(* Logix 5000 project; controller TFF vendor 1 type 14 code 107 rev 33.11; software revision 33.04; part 13 of 38 *)
(* tags used below, declared in another part *)
   AlarmAnalog : AlarmAnalog[50];   // Analog Alarm Array
   AlarmControl : AlarmControl;   // Alarm Control
   AlarmDeviation : AlarmDeviation[20];   // Control Loop Deviation Alarm Array
   AnalogPoint : AnalogInput[50];   // Analog Input Array
   BagInflate : BagInflate;
   CCPSystem : CCPSystem;   // CCP System Data
   ChartMark : ChartMark;   // Chart Mark
   Concentration : Concentration;
   ControlLoop : ControlLoop[20];   // Control Loop Array
   CriteriaFlag : CriteriaFlag;   // Criteria Flag used in CCP Recipe
   DerivedData : DerivedData;   // Derived data (user input and calculated values)
   Diafiltration : Diafiltration;
   DigitalOutput : BOOL[256];   // Digital Output Array these bits are sent to output cards.
   DigitalPoint : DigitalPoint[150];   // Digital Point Array
   Drive : Drive[11];   // Drives Array
   Exchange_OUT : Exchange_OUT;   // Exchange Outputs
   ExternalTCU : BOOL;   // Use of External TCU
   ExternalWeight : BOOL;   // Use of External Weight
   FlowPath : FlowPath[64];   // Flow Path Array
   FQ_Conc : ALIAS FOR Totalizer[0];   // Concentration Totalizer
   FQ_Diaf : ALIAS FOR Totalizer[1];   // DiafiltrationTotalizer
   Gateway : Gateway;   // Gateway Control
   LogVal : LoggedValue;   // Setpoints to be logged
   Membrane_Data : Membrane_Data;   // Membrane Data
   MiscBOOL : BOOL[64];   // Misc BOOL Values
   MiscDINT : DINT[32];   // Misc DINT Values
   MiscREAL : REAL[50];   // Misc Real Values
   Mixer : Mixer;   // Mixer config. structure
   Operation : Operation[6,251];   // Operation Table
   PCV101_Control : PCV_Control;   // PCV101 Control UDT
   PCV201_Control : PCV_Control;   // PCV201 Control UDT
   Phase : Phases[6];   // Phase Control Array
   Prompt : Prompt[7];   // Prompt Array
   PromptTimer : FBD_TIMER;   // Prompt Timer
   SysControl : SysControl;   // General system status and command
   TIC101Control : TCUControl;
   Timers : Timers[22];   // Timer Array
   Totalizer : Totalizers[20];   // Totalizers Array
   UserAlarm : UserAlarm;   // User Alarm (used in CCP Recipe)
   UserTotalizerManagement : UserTotalizerManagement;   // User Totalizer management
   Valve : Valve[100];   // Valve Array

        [2,19].AlarmTimerSP := 2, [2,19].AutoCloseTimer.ACC := 1007, [2,20].Tag := 'XV021', [2,20].CloseStatus := 1, [2,20].ZSOverride := 1, [2,20].EnableCfg := 1, [2,20].StatusWord := 4, [2,20].Status := 4, [2,20].OutputAddress := 52, [2,20].AlarmTimer.PRE := 2000, [2,20].AlarmTimerSP := 2, [2,20].AutoCloseTimer.ACC := 1004, [2,21].Tag := 'XV022', [2,21].Control := 1, [2,21].Auto := 1, [2,21].Manual := 1, [2,21].OpenStatus := 1, [2,21].ZSOverride := 1, [2,21].FailState := 1, [2,21].EnableCfg := 1, [2,21].StatusWord := 2, [2,21].Status := 2, [2,21].OutputAddress := 53, [2,21].AlarmTimer.PRE := 2000, [2,21].AlarmTimerSP := 2, [2,22].Tag := 'XV023', [2,22].CloseStatus := 1, [2,22].ZSOverride := 1, [2,22].EnableCfg := 1, [2,22].StatusWord := 4, [2,22].Status := 4, [2,22].OutputAddress := 54, [2,22].AlarmTimer.PRE := 2000, [2,22].AlarmTimerSP := 2, [2,22].AutoCloseTimer.ACC := 131, [2,23].Tag := 'XV024', [2,23].CloseStatus := 1, [2,23].ZSOverride := 1, [2,23].EnableCfg := 1, [2,23].StatusWord := 4, [2,23].Status := 4, [2,23].OutputAddress := 55, [2,23].AlarmTimer.PRE := 2000, [2,23].AlarmTimerSP := 2, [2,23].AutoCloseTimer.ACC := 1003, [2,24].Tag := 'XV025', [2,24].CloseStatus := 1, [2,24].ZSOverride := 1, [2,24].EnableCfg := 1, [2,24].StatusWord := 4, [2,24].Status := 4, [2,24].OutputAddress := 56, [2,24].AlarmTimer.PRE := 2000, [2,24].AlarmTimerSP := 2, [2,24].AutoCloseTimer.ACC := 1002, [2,25].Tag := 'XV026', [2,25].CloseStatus := 1, [2,25].ZSOverride := 1, [2,25].EnableCfg := 1, [2,25].StatusWord := 4,
        [2,25].Status := 4, [2,25].OutputAddress := 57, [2,25].AlarmTimer.PRE := 2000, [2,25].AlarmTimerSP := 2, [2,25].AutoCloseTimer.ACC := 1002, [2,26].Tag := 'XV028', [2,26].CloseStatus := 1, [2,26].ZSOverride := 1, [2,26].EnableCfg := 1, [2,26].StatusWord := 4, [2,26].Status := 4, [2,26].OutputAddress := 58, [2,26].AlarmTimer.PRE := 2000, [2,26].AlarmTimerSP := 2, [2,26].AutoCloseTimer.ACC := 1002, [2,27].Tag := 'XV029', [2,27].CloseStatus := 1, [2,27].ZSOverride := 1, [2,27].EnableCfg := 1, [2,27].StatusWord := 4, [2,27].Status := 4, [2,27].OutputAddress := 59, [2,27].AlarmTimer.PRE := 2000, [2,27].AlarmTimerSP := 2, [2,28].Tag := 'XV030', [2,28].CloseStatus := 1, [2,28].ZSOverride := 1, [2,28].EnableCfg := 1, [2,28].StatusWord := 4, [2,28].Status := 4, [2,28].OutputAddress := 60, [2,28].AlarmTimer.PRE := 2000, [2,28].AlarmTimerSP := 2, [2,29].Tag := 'XV031', [2,29].Control := 1, [2,29].Auto := 1, [2,29].Manual := 1, [2,29].OpenStatus := 1, [2,29].ZSOverride := 1, [2,29].FailState := 1, [2,29].EnableCfg := 1, [2,29].StatusWord := 2, [2,29].Status := 2, [2,29].OutputAddress := 61, [2,29].AlarmTimer.PRE := 2000, [2,29].AlarmTimerSP := 2, [2,29].AutoCloseTimer.ACC := 1068, [2,30].Tag := 'XV033', [2,30].CloseStatus := 1, [2,30].ZSOverride := 1, [2,30].EnableCfg := 1, [2,30].StatusWord := 4, [2,30].Status := 4, [2,30].OutputAddress := 62, [2,30].AlarmTimer.PRE := 2000, [2,30].AlarmTimerSP := 2, [2,30].AutoCloseTimer.ACC := 1069, [2,31].Tag := 'XV034', [2,31].CloseStatus := 1, [2,31].ZSOverride := 1,
        [2,31].EnableCfg := 1, [2,31].StatusWord := 4, [2,31].Status := 4, [2,31].OutputAddress := 63, [2,31].AlarmTimer.PRE := 2000, [2,31].AlarmTimerSP := 2, [2,31].AutoCloseTimer.ACC := 131, [2,32].CloseStatus := 1, [2,32].PriorityCfg := 1, [2,32].ZSOpenAddress := 32, [2,32].OutputAddress := 68, [2,32].AlarmTimer.PRE := 2000, [2,32].AlarmTimerSP := 2, [2,32].AutoCloseTimer.ACC := 1059, [2,33].OpenStatus := 1, [2,33].PriorityCfg := 1, [2,33].FailState := 1, [2,33].ZSCloseAddress := 33, [2,33].OutputAddress := 69, [2,33].AlarmTimer.PRE := 2000, [2,33].AlarmTimerSP := 2, [2,33].AutoCloseTimer.ACC := 1123, [2,34].OpenStatus := 1, [2,34].PriorityCfg := 1, [2,34].FailState := 1, [2,34].ZSCloseAddress := 34, [2,34].OutputAddress := 70, [2,34].AlarmTimer.PRE := 2000, [2,34].AlarmTimerSP := 2, [2,34].AutoCloseTimer.ACC := 1095, [2,35].OpenStatus := 1, [2,35].PriorityCfg := 1, [2,35].FailState := 1, [2,35].ZSCloseAddress := 35, [2,35].OutputAddress := 71, [2,35].AlarmTimer.PRE := 2000, [2,35].AlarmTimerSP := 2, [2,35].AutoCloseTimer.ACC := 1127, [2,36].OpenStatus := 1, [2,36].PriorityCfg := 1, [2,36].FailState := 1, [2,36].ZSCloseAddress := 36, [2,36].OutputAddress := 72, [2,36].AlarmTimer.PRE := 2000, [2,36].AlarmTimerSP := 2, [2,36].AutoCloseTimer.ACC := 1004, [2,37].CloseStatus := 1, [2,37].PriorityCfg := 1, [2,37].ZSOpenAddress := 37, [2,37].OutputAddress := 73, [2,37].AlarmTimer.PRE := 2000, [2,37].AlarmTimerSP := 2, [2,37].AutoCloseTimer.ACC := 1121, [2,38].CloseStatus := 1, [2,38].Priority := 1, [2,38].PriorityCfg := 1, [2,38].ZSOpenAddress := 38, [2,38].OutputAddress := 40, [2,38].AlarmTimer.PRE := 2000, [2,38].AlarmTimerSP := 2,
        [2,38].AutoCloseTimer.ACC := 1135, [2,39].CloseStatus := 1, [2,39].Priority := 1, [2,39].PriorityCfg := 1, [2,39].ZSOpenAddress := 39, [2,39].OutputAddress := 41, [2,39].AlarmTimer.PRE := 2000, [2,39].AlarmTimerSP := 2, [2,39].AutoCloseTimer.ACC := 1121, [2,40].CloseStatus := 1, [2,40].Priority := 1, [2,40].PriorityCfg := 1, [2,40].ZSOpenAddress := 40, [2,40].OutputAddress := 42, [2,40].AlarmTimer.PRE := 2000, [2,40].AlarmTimerSP := 2, [2,40].AutoCloseTimer.ACC := 1112, [2,41].CloseStatus := 1, [2,41].Priority := 1, [2,41].PriorityCfg := 1, [2,41].ZSOpenAddress := 41, [2,41].OutputAddress := 43, [2,41].AlarmTimer.PRE := 2000, [2,41].AlarmTimerSP := 2, [2,42].CloseStatus := 1, [2,42].Priority := 1, [2,42].PriorityCfg := 1, [2,42].ZSOpenAddress := 42, [2,42].OutputAddress := 44, [2,42].AlarmTimer.PRE := 2000, [2,42].AlarmTimerSP := 2, [2,43].CloseStatus := 1, [2,43].Priority := 1, [2,43].PriorityCfg := 1, [2,43].ZSOpenAddress := 43, [2,43].OutputAddress := 52, [2,43].AlarmTimer.PRE := 2000, [2,43].AlarmTimerSP := 2, [2,44].CloseStatus := 1, [2,44].Priority := 1, [2,44].PriorityCfg := 1, [2,44].ZSOpenAddress := 44, [2,44].OutputAddress := 53, [2,44].AlarmTimer.PRE := 2000, [2,44].AlarmTimerSP := 2, [2,45].CloseStatus := 1, [2,45].Priority := 1, [2,45].PriorityCfg := 1, [2,45].ZSOpenAddress := 45, [2,45].OutputAddress := 54, [2,45].AlarmTimer.PRE := 2000, [2,45].AlarmTimerSP := 2, [2,46].CloseStatus := 1, [2,46].Priority := 1, [2,46].PriorityCfg := 1, [2,46].ZSOpenAddress := 46, [2,46].OutputAddress := 55, [2,46].AlarmTimer.PRE := 2000, [2,46].AlarmTimerSP := 2, [2,47].OpenStatus := 1,
        [2,47].Priority := 1, [2,47].PriorityCfg := 1, [2,47].FailState := 1, [2,47].ZSCloseAddress := 47, [2,47].OutputAddress := 45, [2,47].AlarmTimer.PRE := 2000, [2,47].AlarmTimerSP := 2, [2,48].FailState := 1, [2,48].ZSCloseAddress := 48, [2,48].OutputAddress := 80, [2,49].FailState := 1, [2,49].ZSCloseAddress := 49, [2,49].OutputAddress := 81, [2,50].FailState := 1, [2,50].ZSCloseAddress := 50, [2,50].OutputAddress := 82, [2,51].OpenStatus := 1, [2,51].FailState := 1, [2,51].ZSCloseAddress := 51, [2,51].OutputAddress := 83, [2,52].OpenStatus := 1, [2,52].FailState := 1, [2,52].ZSCloseAddress := 52, [2,52].OutputAddress := 84, [2,53].CloseStatus := 1, [2,53].FailState := 1, [2,53].ZSCloseAddress := 53, [2,53].OutputAddress := 85, [2,54].CloseStatus := 1, [2,54].FailState := 1, [2,54].ZSCloseAddress := 54, [2,54].OutputAddress := 86, [2,55].CloseStatus := 1, [2,55].FailState := 1, [2,55].ZSCloseAddress := 55, [2,55].OutputAddress := 87, [2,56].CloseStatus := 1, [2,58].CloseStatus := 1, [2,59].CloseStatus := 1, [3,0].CloseStatus := 1, [3,0].EnableCfg := 1, [3,0].StatusWord := 4, [3,0].Status := 4, [3,0].OutputAddress := 32, [3,1].CloseStatus := 1, [3,1].EnableCfg := 1, [3,1].StatusWord := 4, [3,1].Status := 4, [3,1].OutputAddress := 33, [3,2].CloseStatus := 1, [3,2].EnableCfg := 1, [3,2].StatusWord := 4, [3,2].Status := 4, [3,2].OutputAddress := 34, [3,3].CloseStatus := 1, [3,3].EnableCfg := 1, [3,3].StatusWord := 4, [3,3].Status := 4, [3,3].OutputAddress := 35, [3,4].CloseStatus := 1,
        [3,4].EnableCfg := 1, [3,4].StatusWord := 4, [3,4].Status := 4, [3,4].OutputAddress := 36, [3,5].CloseStatus := 1, [3,5].EnableCfg := 1, [3,5].StatusWord := 4, [3,5].Status := 4, [3,5].OutputAddress := 37, [3,6].CloseStatus := 1, [3,6].EnableCfg := 1, [3,6].StatusWord := 4, [3,6].Status := 4, [3,6].OutputAddress := 38, [3,7].CloseStatus := 1, [3,7].EnableCfg := 1, [3,7].StatusWord := 4, [3,7].Status := 4, [3,7].OutputAddress := 39, [3,8].CloseStatus := 1, [3,8].EnableCfg := 1, [3,8].StatusWord := 4, [3,8].Status := 4, [3,8].OutputAddress := 40, [3,9].CloseStatus := 1, [3,9].EnableCfg := 1, [3,9].StatusWord := 4, [3,9].Status := 4, [3,9].OutputAddress := 41, [3,10].CloseStatus := 1, [3,10].EnableCfg := 1, [3,10].StatusWord := 4, [3,10].Status := 4, [3,10].OutputAddress := 42, [3,11].CloseStatus := 1, [3,11].FailState := 1, [3,11].EnableCfg := 1, [3,11].StatusWord := 4, [3,11].Status := 4, [3,11].OutputAddress := 43, [3,12].CloseStatus := 1, [3,12].FailState := 1, [3,12].EnableCfg := 1, [3,12].StatusWord := 4, [3,12].Status := 4, [3,12].OutputAddress := 44, [3,13].CloseStatus := 1, [3,13].FailState := 1, [3,13].EnableCfg := 1, [3,13].StatusWord := 4, [3,13].Status := 4, [3,13].OutputAddress := 45, [3,14].CloseStatus := 1, [3,14].EnableCfg := 1, [3,14].StatusWord := 4, [3,14].Status := 4, [3,14].OutputAddress := 46, [3,15].CloseStatus := 1, [3,15].FailState := 1, [3,15].EnableCfg := 1,
        [3,15].StatusWord := 4, [3,15].Status := 4, [3,15].OutputAddress := 47, [3,16].CloseStatus := 1, [3,16].EnableCfg := 1, [3,16].StatusWord := 4, [3,16].Status := 4, [3,16].OutputAddress := 48, [3,17].CloseStatus := 1, [3,17].FailState := 1, [3,17].EnableCfg := 1, [3,17].StatusWord := 4, [3,17].Status := 4, [3,17].OutputAddress := 49, [3,18].CloseStatus := 1, [3,18].EnableCfg := 1, [3,18].StatusWord := 4, [3,18].Status := 4, [3,18].OutputAddress := 50, [3,19].CloseStatus := 1, [3,19].EnableCfg := 1, [3,19].StatusWord := 4, [3,19].Status := 4, [3,19].OutputAddress := 51, [3,20].CloseStatus := 1, [3,20].EnableCfg := 1, [3,20].StatusWord := 4, [3,20].Status := 4, [3,20].OutputAddress := 52, [3,21].CloseStatus := 1, [3,21].FailState := 1, [3,21].EnableCfg := 1, [3,21].StatusWord := 4, [3,21].Status := 4, [3,21].OutputAddress := 53, [3,22].CloseStatus := 1, [3,22].EnableCfg := 1, [3,22].StatusWord := 4, [3,22].Status := 4, [3,22].OutputAddress := 54, [3,23].CloseStatus := 1, [3,23].EnableCfg := 1, [3,23].StatusWord := 4, [3,23].Status := 4, [3,23].OutputAddress := 55, [3,24].CloseStatus := 1, [3,24].EnableCfg := 1, [3,24].StatusWord := 4, [3,24].Status := 4, [3,24].OutputAddress := 56, [3,25].CloseStatus := 1, [3,25].EnableCfg := 1, [3,25].StatusWord := 4, [3,25].Status := 4, [3,25].OutputAddress := 57, [3,26].CloseStatus := 1, [3,26].EnableCfg := 1, [3,26].StatusWord := 4, [3,26].Status := 4, [3,26].OutputAddress := 58,
        [3,27].CloseStatus := 1, [3,27].EnableCfg := 1, [3,27].StatusWord := 4, [3,27].Status := 4, [3,27].OutputAddress := 59, [3,28].CloseStatus := 1, [3,28].EnableCfg := 1, [3,28].StatusWord := 4, [3,28].Status := 4, [3,28].OutputAddress := 60, [3,29].CloseStatus := 1, [3,29].FailState := 1, [3,29].EnableCfg := 1, [3,29].StatusWord := 4, [3,29].Status := 4, [3,29].OutputAddress := 61, [3,30].CloseStatus := 1, [3,30].EnableCfg := 1, [3,30].StatusWord := 4, [3,30].Status := 4, [3,30].OutputAddress := 62, [3,31].CloseStatus := 1, [3,31].EnableCfg := 1, [3,31].StatusWord := 4, [3,31].Status := 4, [3,31].OutputAddress := 63, [4,0].Tag := 'XV001', [4,0].CloseStatus := 1, [4,0].ZSOverride := 1, [4,0].EnableCfg := 1, [4,0].StatusWord := 4, [4,0].Status := 4, [4,0].OutputAddress := 32, [4,0].AlarmTimer.PRE := 2000, [4,0].AlarmTimerSP := 2, [4,1].Tag := 'XV002', [4,1].CloseStatus := 1, [4,1].ZSOverride := 1, [4,1].EnableCfg := 1, [4,1].StatusWord := 4, [4,1].Status := 4, [4,1].OutputAddress := 33, [4,1].AlarmTimer.PRE := 2000, [4,1].AlarmTimerSP := 2, [4,1].AutoCloseTimer.ACC := 1103, [4,2].Tag := 'XV003', [4,2].CloseStatus := 1, [4,2].ZSOverride := 1, [4,2].EnableCfg := 1, [4,2].StatusWord := 4, [4,2].Status := 4, [4,2].OutputAddress := 34, [4,2].AlarmTimer.PRE := 2000, [4,2].AlarmTimerSP := 2, [4,2].AutoCloseTimer.ACC := 1032, [4,3].Tag := 'XV004', [4,3].CloseStatus := 1, [4,3].ZSOverride := 1, [4,3].EnableCfg := 1, [4,3].StatusWord := 4,
        [4,3].Status := 4, [4,3].OutputAddress := 35, [4,3].AlarmTimer.PRE := 2000, [4,3].AlarmTimerSP := 2, [4,3].AutoCloseTimer.ACC := 1115, [4,4].Tag := 'XV005', [4,4].CloseStatus := 1, [4,4].ZSOverride := 1, [4,4].EnableCfg := 1, [4,4].StatusWord := 4, [4,4].Status := 4, [4,4].OutputAddress := 36, [4,4].AlarmTimer.PRE := 2000, [4,4].AlarmTimerSP := 2, [4,4].AutoCloseTimer.ACC := 1104, [4,5].Tag := 'XV006', [4,5].CloseStatus := 1, [4,5].ZSOverride := 1, [4,5].EnableCfg := 1, [4,5].StatusWord := 4, [4,5].Status := 4, [4,5].OutputAddress := 37, [4,5].AlarmTimer.PRE := 2000, [4,5].AlarmTimerSP := 2, [4,5].AutoCloseTimer.ACC := 1104, [4,6].Tag := 'XV007', [4,6].CloseStatus := 1, [4,6].ZSOverride := 1, [4,6].EnableCfg := 1, [4,6].StatusWord := 4, [4,6].Status := 4, [4,6].OutputAddress := 38, [4,6].AlarmTimer.PRE := 2000, [4,6].AlarmTimerSP := 2, [4,6].AutoCloseTimer.ACC := 1104, [4,7].Tag := 'XV008', [4,7].CloseStatus := 1, [4,7].ZSOverride := 1, [4,7].EnableCfg := 1, [4,7].StatusWord := 4, [4,7].Status := 4, [4,7].OutputAddress := 39, [4,7].AlarmTimer.PRE := 2000, [4,7].AlarmTimerSP := 2, [4,7].AutoCloseTimer.ACC := 1104, [4,8].Tag := 'XV009', [4,8].CloseStatus := 1, [4,8].ZSOverride := 1, [4,8].EnableCfg := 1, [4,8].StatusWord := 4, [4,8].Status := 4, [4,8].OutputAddress := 40, [4,8].AlarmTimer.PRE := 2000, [4,8].AlarmTimerSP := 2, [4,8].AutoCloseTimer.ACC := 1104, [4,9].Tag := 'XV010', [4,9].CloseStatus := 1, [4,9].ZSOverride := 1, [4,9].EnableCfg := 1, [4,9].StatusWord := 4,
        [4,9].Status := 4, [4,9].OutputAddress := 41, [4,9].AlarmTimer.PRE := 2000, [4,9].AlarmTimerSP := 2, [4,9].AutoCloseTimer.ACC := 1105, [4,10].Tag := 'XV011', [4,10].CloseStatus := 1, [4,10].ZSOverride := 1, [4,10].EnableCfg := 1, [4,10].StatusWord := 4, [4,10].Status := 4, [4,10].OutputAddress := 42, [4,10].AlarmTimer.PRE := 2000, [4,10].AlarmTimerSP := 2, [4,10].AutoCloseTimer.ACC := 1104, [4,11].Tag := 'XV012', [4,11].Control := 1, [4,11].Auto := 1, [4,11].Manual := 1, [4,11].OpenStatus := 1, [4,11].ZSOverride := 1, [4,11].FailState := 1, [4,11].EnableCfg := 1, [4,11].StatusWord := 2, [4,11].Status := 2, [4,11].OutputAddress := 43, [4,11].AlarmTimer.PRE := 2000, [4,11].AlarmTimerSP := 2, [4,11].AutoCloseTimer.ACC := 1103, [4,12].Tag := 'XV013', [4,12].Control := 1, [4,12].Auto := 1, [4,12].Manual := 1, [4,12].OpenStatus := 1, [4,12].ZSOverride := 1, [4,12].FailState := 1, [4,12].EnableCfg := 1, [4,12].StatusWord := 2, [4,12].Status := 2, [4,12].OutputAddress := 44, [4,12].AlarmTimer.PRE := 2000, [4,12].AlarmTimerSP := 2, [4,12].AutoCloseTimer.ACC := 1072, [4,13].Tag := 'XV014', [4,13].Control := 1, [4,13].Auto := 1, [4,13].Manual := 1, [4,13].OpenStatus := 1, [4,13].ZSOverride := 1, [4,13].FailState := 1, [4,13].EnableCfg := 1, [4,13].StatusWord := 2, [4,13].Status := 2, [4,13].OutputAddress := 45, [4,13].AlarmTimer.PRE := 2000, [4,13].AlarmTimerSP := 2, [4,13].AutoCloseTimer.ACC := 1016, [4,14].Tag := 'XV015', [4,14].CloseStatus := 1, [4,14].ZSOverride := 1,
        [4,14].EnableCfg := 1, [4,14].StatusWord := 4, [4,14].Status := 4, [4,14].OutputAddress := 46, [4,14].AlarmTimer.PRE := 2000, [4,14].AlarmTimerSP := 2, [4,15].Tag := 'XV016', [4,15].Control := 1, [4,15].Auto := 1, [4,15].Manual := 1, [4,15].OpenStatus := 1, [4,15].ZSOverride := 1, [4,15].FailState := 1, [4,15].EnableCfg := 1, [4,15].StatusWord := 2, [4,15].Status := 2, [4,15].OutputAddress := 47, [4,15].AlarmTimer.PRE := 2000, [4,15].AlarmTimerSP := 2, [4,16].Tag := 'XV017', [4,16].CloseStatus := 1, [4,16].ZSOverride := 1, [4,16].EnableCfg := 1, [4,16].StatusWord := 4, [4,16].Status := 4, [4,16].OutputAddress := 48, [4,16].AlarmTimer.PRE := 2000, [4,16].AlarmTimerSP := 2, [4,17].Tag := 'XV018', [4,17].Control := 1, [4,17].Auto := 1, [4,17].Manual := 1, [4,17].OpenStatus := 1, [4,17].ZSOverride := 1, [4,17].FailState := 1, [4,17].EnableCfg := 1, [4,17].StatusWord := 2, [4,17].Status := 2, [4,17].OutputAddress := 49, [4,17].AlarmTimer.PRE := 2000, [4,17].AlarmTimerSP := 2, [4,17].AutoCloseTimer.ACC := 1594, [4,18].Tag := 'XV019', [4,18].CloseStatus := 1, [4,18].ZSOverride := 1, [4,18].EnableCfg := 1, [4,18].StatusWord := 4, [4,18].Status := 4, [4,18].OutputAddress := 50, [4,18].AlarmTimer.PRE := 2000, [4,18].AlarmTimerSP := 2, [4,18].AutoCloseTimer.ACC := 137, [4,19].Tag := 'XV020', [4,19].CloseStatus := 1, [4,19].ZSOverride := 1, [4,19].EnableCfg := 1, [4,19].StatusWord := 4, [4,19].Status := 4, [4,19].OutputAddress := 51, [4,19].AlarmTimer.PRE := 2000,
        [4,19].AlarmTimerSP := 2, [4,19].AutoCloseTimer.ACC := 1007, [4,20].Tag := 'XV021', [4,20].CloseStatus := 1, [4,20].ZSOverride := 1, [4,20].EnableCfg := 1, [4,20].StatusWord := 4, [4,20].Status := 4, [4,20].OutputAddress := 52, [4,20].AlarmTimer.PRE := 2000, [4,20].AlarmTimerSP := 2, [4,20].AutoCloseTimer.ACC := 1004, [4,21].Tag := 'XV022', [4,21].Control := 1, [4,21].Auto := 1, [4,21].Manual := 1, [4,21].OpenStatus := 1, [4,21].ZSOverride := 1, [4,21].FailState := 1, [4,21].EnableCfg := 1, [4,21].StatusWord := 2, [4,21].Status := 2, [4,21].OutputAddress := 53, [4,21].AlarmTimer.PRE := 2000, [4,21].AlarmTimerSP := 2, [4,22].Tag := 'XV023', [4,22].CloseStatus := 1, [4,22].ZSOverride := 1, [4,22].EnableCfg := 1, [4,22].StatusWord := 4, [4,22].Status := 4, [4,22].OutputAddress := 54, [4,22].AlarmTimer.PRE := 2000, [4,22].AlarmTimerSP := 2, [4,22].AutoCloseTimer.ACC := 131, [4,23].Tag := 'XV024', [4,23].CloseStatus := 1, [4,23].ZSOverride := 1, [4,23].EnableCfg := 1, [4,23].StatusWord := 4, [4,23].Status := 4, [4,23].OutputAddress := 55, [4,23].AlarmTimer.PRE := 2000, [4,23].AlarmTimerSP := 2, [4,23].AutoCloseTimer.ACC := 1003, [4,24].Tag := 'XV025', [4,24].CloseStatus := 1, [4,24].ZSOverride := 1, [4,24].EnableCfg := 1, [4,24].StatusWord := 4, [4,24].Status := 4, [4,24].OutputAddress := 56, [4,24].AlarmTimer.PRE := 2000, [4,24].AlarmTimerSP := 2, [4,24].AutoCloseTimer.ACC := 1002, [4,25].Tag := 'XV026', [4,25].CloseStatus := 1, [4,25].ZSOverride := 1, [4,25].EnableCfg := 1, [4,25].StatusWord := 4,
        [4,25].Status := 4, [4,25].OutputAddress := 57, [4,25].AlarmTimer.PRE := 2000, [4,25].AlarmTimerSP := 2, [4,25].AutoCloseTimer.ACC := 1002, [4,26].Tag := 'XV028', [4,26].CloseStatus := 1, [4,26].ZSOverride := 1, [4,26].EnableCfg := 1, [4,26].StatusWord := 4, [4,26].Status := 4, [4,26].OutputAddress := 58, [4,26].AlarmTimer.PRE := 2000, [4,26].AlarmTimerSP := 2, [4,26].AutoCloseTimer.ACC := 1002, [4,27].Tag := 'XV029', [4,27].CloseStatus := 1, [4,27].ZSOverride := 1, [4,27].EnableCfg := 1, [4,27].StatusWord := 4, [4,27].Status := 4, [4,27].OutputAddress := 59, [4,27].AlarmTimer.PRE := 2000, [4,27].AlarmTimerSP := 2, [4,28].Tag := 'XV030', [4,28].CloseStatus := 1, [4,28].ZSOverride := 1, [4,28].EnableCfg := 1, [4,28].StatusWord := 4, [4,28].Status := 4, [4,28].OutputAddress := 60, [4,28].AlarmTimer.PRE := 2000, [4,28].AlarmTimerSP := 2, [4,29].Tag := 'XV031', [4,29].Control := 1, [4,29].Auto := 1, [4,29].Manual := 1, [4,29].OpenStatus := 1, [4,29].ZSOverride := 1, [4,29].FailState := 1, [4,29].EnableCfg := 1, [4,29].StatusWord := 2, [4,29].Status := 2, [4,29].OutputAddress := 61, [4,29].AlarmTimer.PRE := 2000, [4,29].AlarmTimerSP := 2, [4,29].AutoCloseTimer.ACC := 1068, [4,30].Tag := 'XV033', [4,30].CloseStatus := 1, [4,30].ZSOverride := 1, [4,30].EnableCfg := 1, [4,30].StatusWord := 4, [4,30].Status := 4, [4,30].OutputAddress := 62, [4,30].AlarmTimer.PRE := 2000, [4,30].AlarmTimerSP := 2, [4,30].AutoCloseTimer.ACC := 1069, [4,31].Tag := 'XV034', [4,31].CloseStatus := 1, [4,31].ZSOverride := 1,
        [4,31].EnableCfg := 1, [4,31].StatusWord := 4, [4,31].Status := 4, [4,31].OutputAddress := 63, [4,31].AlarmTimer.PRE := 2000, [4,31].AlarmTimerSP := 2, [4,31].AutoCloseTimer.ACC := 131, [4,32].CloseStatus := 1, [4,32].PriorityCfg := 1, [4,32].ZSOpenAddress := 32, [4,32].OutputAddress := 68, [4,32].AlarmTimer.PRE := 2000, [4,32].AlarmTimerSP := 2, [4,32].AutoCloseTimer.ACC := 1059, [4,33].OpenStatus := 1, [4,33].PriorityCfg := 1, [4,33].FailState := 1, [4,33].ZSCloseAddress := 33, [4,33].OutputAddress := 69, [4,33].AlarmTimer.PRE := 2000, [4,33].AlarmTimerSP := 2, [4,33].AutoCloseTimer.ACC := 1123, [4,34].OpenStatus := 1, [4,34].PriorityCfg := 1, [4,34].FailState := 1, [4,34].ZSCloseAddress := 34, [4,34].OutputAddress := 70, [4,34].AlarmTimer.PRE := 2000, [4,34].AlarmTimerSP := 2, [4,34].AutoCloseTimer.ACC := 1095, [4,35].OpenStatus := 1, [4,35].PriorityCfg := 1, [4,35].FailState := 1, [4,35].ZSCloseAddress := 35, [4,35].OutputAddress := 71, [4,35].AlarmTimer.PRE := 2000, [4,35].AlarmTimerSP := 2, [4,35].AutoCloseTimer.ACC := 1127, [4,36].OpenStatus := 1, [4,36].PriorityCfg := 1, [4,36].FailState := 1, [4,36].ZSCloseAddress := 36, [4,36].OutputAddress := 72, [4,36].AlarmTimer.PRE := 2000, [4,36].AlarmTimerSP := 2, [4,36].AutoCloseTimer.ACC := 1004, [4,37].CloseStatus := 1, [4,37].PriorityCfg := 1, [4,37].ZSOpenAddress := 37, [4,37].OutputAddress := 73, [4,37].AlarmTimer.PRE := 2000, [4,37].AlarmTimerSP := 2, [4,37].AutoCloseTimer.ACC := 1121, [4,38].CloseStatus := 1, [4,38].Priority := 1, [4,38].PriorityCfg := 1, [4,38].ZSOpenAddress := 38, [4,38].OutputAddress := 40, [4,38].AlarmTimer.PRE := 2000, [4,38].AlarmTimerSP := 2,
        [4,38].AutoCloseTimer.ACC := 1135, [4,39].CloseStatus := 1, [4,39].Priority := 1, [4,39].PriorityCfg := 1, [4,39].ZSOpenAddress := 39, [4,39].OutputAddress := 41, [4,39].AlarmTimer.PRE := 2000, [4,39].AlarmTimerSP := 2, [4,39].AutoCloseTimer.ACC := 1121, [4,40].CloseStatus := 1, [4,40].Priority := 1, [4,40].PriorityCfg := 1, [4,40].ZSOpenAddress := 40, [4,40].OutputAddress := 42, [4,40].AlarmTimer.PRE := 2000, [4,40].AlarmTimerSP := 2, [4,40].AutoCloseTimer.ACC := 1112, [4,41].CloseStatus := 1, [4,41].Priority := 1, [4,41].PriorityCfg := 1, [4,41].ZSOpenAddress := 41, [4,41].OutputAddress := 43, [4,41].AlarmTimer.PRE := 2000, [4,41].AlarmTimerSP := 2, [4,42].CloseStatus := 1, [4,42].Priority := 1, [4,42].PriorityCfg := 1, [4,42].ZSOpenAddress := 42, [4,42].OutputAddress := 44, [4,42].AlarmTimer.PRE := 2000, [4,42].AlarmTimerSP := 2, [4,43].CloseStatus := 1, [4,43].Priority := 1, [4,43].PriorityCfg := 1, [4,43].ZSOpenAddress := 43, [4,43].OutputAddress := 52, [4,43].AlarmTimer.PRE := 2000, [4,43].AlarmTimerSP := 2, [4,44].CloseStatus := 1, [4,44].Priority := 1, [4,44].PriorityCfg := 1, [4,44].ZSOpenAddress := 44, [4,44].OutputAddress := 53, [4,44].AlarmTimer.PRE := 2000, [4,44].AlarmTimerSP := 2, [4,45].CloseStatus := 1, [4,45].Priority := 1, [4,45].PriorityCfg := 1, [4,45].ZSOpenAddress := 45, [4,45].OutputAddress := 54, [4,45].AlarmTimer.PRE := 2000, [4,45].AlarmTimerSP := 2, [4,46].CloseStatus := 1, [4,46].Priority := 1, [4,46].PriorityCfg := 1, [4,46].ZSOpenAddress := 46, [4,46].OutputAddress := 55, [4,46].AlarmTimer.PRE := 2000, [4,46].AlarmTimerSP := 2, [4,47].OpenStatus := 1,
        [4,47].Priority := 1, [4,47].PriorityCfg := 1, [4,47].FailState := 1, [4,47].ZSCloseAddress := 47, [4,47].OutputAddress := 45, [4,47].AlarmTimer.PRE := 2000, [4,47].AlarmTimerSP := 2, [4,48].FailState := 1, [4,48].ZSCloseAddress := 48, [4,48].OutputAddress := 80, [4,49].FailState := 1, [4,49].ZSCloseAddress := 49, [4,49].OutputAddress := 81, [4,50].FailState := 1, [4,50].ZSCloseAddress := 50, [4,50].OutputAddress := 82, [4,51].OpenStatus := 1, [4,51].FailState := 1, [4,51].ZSCloseAddress := 51, [4,51].OutputAddress := 83, [4,52].OpenStatus := 1, [4,52].FailState := 1, [4,52].ZSCloseAddress := 52, [4,52].OutputAddress := 84, [4,53].CloseStatus := 1, [4,53].FailState := 1, [4,53].ZSCloseAddress := 53, [4,53].OutputAddress := 85, [4,54].CloseStatus := 1, [4,54].FailState := 1, [4,54].ZSCloseAddress := 54, [4,54].OutputAddress := 86, [4,55].CloseStatus := 1, [4,55].FailState := 1, [4,55].ZSCloseAddress := 55, [4,55].OutputAddress := 87, [4,56].CloseStatus := 1, [4,58].CloseStatus := 1, [4,59].CloseStatus := 1, [5,0].Tag := 'XV001', [5,0].CloseStatus := 1, [5,0].ZSOverride := 1, [5,0].EnableCfg := 1, [5,0].StatusWord := 4, [5,0].Status := 4, [5,0].OutputAddress := 32, [5,0].AlarmTimer.PRE := 2000, [5,0].AlarmTimerSP := 2, [5,1].Tag := 'XV002', [5,1].CloseStatus := 1, [5,1].ZSOverride := 1, [5,1].EnableCfg := 1, [5,1].StatusWord := 4, [5,1].Status := 4, [5,1].OutputAddress := 33, [5,1].AlarmTimer.PRE := 2000, [5,1].AlarmTimerSP := 2, [5,1].AutoCloseTimer.ACC := 1103, [5,2].Tag := 'XV003', [5,2].CloseStatus := 1,
        [5,2].ZSOverride := 1, [5,2].EnableCfg := 1, [5,2].StatusWord := 4, [5,2].Status := 4, [5,2].OutputAddress := 34, [5,2].AlarmTimer.PRE := 2000, [5,2].AlarmTimerSP := 2, [5,2].AutoCloseTimer.ACC := 1032, [5,3].Tag := 'XV004', [5,3].CloseStatus := 1, [5,3].ZSOverride := 1, [5,3].EnableCfg := 1, [5,3].StatusWord := 4, [5,3].Status := 4, [5,3].OutputAddress := 35, [5,3].AlarmTimer.PRE := 2000, [5,3].AlarmTimerSP := 2, [5,3].AutoCloseTimer.ACC := 1115, [5,4].Tag := 'XV005', [5,4].CloseStatus := 1, [5,4].ZSOverride := 1, [5,4].EnableCfg := 1, [5,4].StatusWord := 4, [5,4].Status := 4, [5,4].OutputAddress := 36, [5,4].AlarmTimer.PRE := 2000, [5,4].AlarmTimerSP := 2, [5,4].AutoCloseTimer.ACC := 1104, [5,5].Tag := 'XV006', [5,5].CloseStatus := 1, [5,5].ZSOverride := 1, [5,5].EnableCfg := 1, [5,5].StatusWord := 4, [5,5].Status := 4, [5,5].OutputAddress := 37, [5,5].AlarmTimer.PRE := 2000, [5,5].AlarmTimerSP := 2, [5,5].AutoCloseTimer.ACC := 1104, [5,6].Tag := 'XV007', [5,6].CloseStatus := 1, [5,6].ZSOverride := 1, [5,6].EnableCfg := 1, [5,6].StatusWord := 4, [5,6].Status := 4, [5,6].OutputAddress := 38, [5,6].AlarmTimer.PRE := 2000, [5,6].AlarmTimerSP := 2, [5,6].AutoCloseTimer.ACC := 1104, [5,7].Tag := 'XV008', [5,7].CloseStatus := 1, [5,7].ZSOverride := 1, [5,7].EnableCfg := 1, [5,7].StatusWord := 4, [5,7].Status := 4, [5,7].OutputAddress := 39, [5,7].AlarmTimer.PRE := 2000, [5,7].AlarmTimerSP := 2, [5,7].AutoCloseTimer.ACC := 1104, [5,8].Tag := 'XV009', [5,8].CloseStatus := 1,
        [5,8].ZSOverride := 1, [5,8].EnableCfg := 1, [5,8].StatusWord := 4, [5,8].Status := 4, [5,8].OutputAddress := 40, [5,8].AlarmTimer.PRE := 2000, [5,8].AlarmTimerSP := 2, [5,8].AutoCloseTimer.ACC := 1104, [5,9].Tag := 'XV010', [5,9].CloseStatus := 1, [5,9].ZSOverride := 1, [5,9].EnableCfg := 1, [5,9].StatusWord := 4, [5,9].Status := 4, [5,9].OutputAddress := 41, [5,9].AlarmTimer.PRE := 2000, [5,9].AlarmTimerSP := 2, [5,9].AutoCloseTimer.ACC := 1105, [5,10].Tag := 'XV011', [5,10].CloseStatus := 1, [5,10].ZSOverride := 1, [5,10].EnableCfg := 1, [5,10].StatusWord := 4, [5,10].Status := 4, [5,10].OutputAddress := 42, [5,10].AlarmTimer.PRE := 2000, [5,10].AlarmTimerSP := 2, [5,10].AutoCloseTimer.ACC := 1104, [5,11].Tag := 'XV012', [5,11].Control := 1, [5,11].Auto := 1, [5,11].Manual := 1, [5,11].OpenStatus := 1, [5,11].ZSOverride := 1, [5,11].FailState := 1, [5,11].EnableCfg := 1, [5,11].StatusWord := 2, [5,11].Status := 2, [5,11].OutputAddress := 43, [5,11].AlarmTimer.PRE := 2000, [5,11].AlarmTimerSP := 2, [5,11].AutoCloseTimer.ACC := 1103, [5,12].Tag := 'XV013', [5,12].Control := 1, [5,12].Auto := 1, [5,12].Manual := 1, [5,12].OpenStatus := 1, [5,12].ZSOverride := 1, [5,12].FailState := 1, [5,12].EnableCfg := 1, [5,12].StatusWord := 2, [5,12].Status := 2, [5,12].OutputAddress := 44, [5,12].AlarmTimer.PRE := 2000, [5,12].AlarmTimerSP := 2, [5,12].AutoCloseTimer.ACC := 1072, [5,13].Tag := 'XV014', [5,13].Control := 1, [5,13].Auto := 1, [5,13].Manual := 1,
        [5,13].OpenStatus := 1, [5,13].ZSOverride := 1, [5,13].FailState := 1, [5,13].EnableCfg := 1, [5,13].StatusWord := 2, [5,13].Status := 2, [5,13].OutputAddress := 45, [5,13].AlarmTimer.PRE := 2000, [5,13].AlarmTimerSP := 2, [5,13].AutoCloseTimer.ACC := 1016, [5,14].Tag := 'XV015', [5,14].CloseStatus := 1, [5,14].ZSOverride := 1, [5,14].EnableCfg := 1, [5,14].StatusWord := 4, [5,14].Status := 4, [5,14].OutputAddress := 46, [5,14].AlarmTimer.PRE := 2000, [5,14].AlarmTimerSP := 2, [5,15].Tag := 'XV016', [5,15].Control := 1, [5,15].Auto := 1, [5,15].Manual := 1, [5,15].OpenStatus := 1, [5,15].ZSOverride := 1, [5,15].FailState := 1, [5,15].EnableCfg := 1, [5,15].StatusWord := 2, [5,15].Status := 2, [5,15].OutputAddress := 47, [5,15].AlarmTimer.PRE := 2000, [5,15].AlarmTimerSP := 2, [5,16].Tag := 'XV017', [5,16].CloseStatus := 1, [5,16].ZSOverride := 1, [5,16].EnableCfg := 1, [5,16].StatusWord := 4, [5,16].Status := 4, [5,16].OutputAddress := 48, [5,16].AlarmTimer.PRE := 2000, [5,16].AlarmTimerSP := 2, [5,17].Tag := 'XV018', [5,17].Control := 1, [5,17].Auto := 1, [5,17].Manual := 1, [5,17].OpenStatus := 1, [5,17].ZSOverride := 1, [5,17].FailState := 1, [5,17].EnableCfg := 1, [5,17].StatusWord := 2, [5,17].Status := 2, [5,17].OutputAddress := 49, [5,17].AlarmTimer.PRE := 2000, [5,17].AlarmTimerSP := 2, [5,17].AutoCloseTimer.ACC := 1594, [5,18].Tag := 'XV019', [5,18].CloseStatus := 1, [5,18].ZSOverride := 1, [5,18].EnableCfg := 1, [5,18].StatusWord := 4,
        [5,18].Status := 4, [5,18].OutputAddress := 50, [5,18].AlarmTimer.PRE := 2000, [5,18].AlarmTimerSP := 2, [5,18].AutoCloseTimer.ACC := 137, [5,19].Tag := 'XV020', [5,19].CloseStatus := 1, [5,19].ZSOverride := 1, [5,19].EnableCfg := 1, [5,19].StatusWord := 4, [5,19].Status := 4, [5,19].OutputAddress := 51, [5,19].AlarmTimer.PRE := 2000, [5,19].AlarmTimerSP := 2, [5,19].AutoCloseTimer.ACC := 1007, [5,20].Tag := 'XV021', [5,20].CloseStatus := 1, [5,20].ZSOverride := 1, [5,20].EnableCfg := 1, [5,20].StatusWord := 4, [5,20].Status := 4, [5,20].OutputAddress := 52, [5,20].AlarmTimer.PRE := 2000, [5,20].AlarmTimerSP := 2, [5,20].AutoCloseTimer.ACC := 1004, [5,21].Tag := 'XV022', [5,21].Control := 1, [5,21].Auto := 1, [5,21].Manual := 1, [5,21].OpenStatus := 1, [5,21].ZSOverride := 1, [5,21].FailState := 1, [5,21].EnableCfg := 1, [5,21].StatusWord := 2, [5,21].Status := 2, [5,21].OutputAddress := 53, [5,21].AlarmTimer.PRE := 2000, [5,21].AlarmTimerSP := 2, [5,22].Tag := 'XV023', [5,22].CloseStatus := 1, [5,22].ZSOverride := 1, [5,22].EnableCfg := 1, [5,22].StatusWord := 4, [5,22].Status := 4, [5,22].OutputAddress := 54, [5,22].AlarmTimer.PRE := 2000, [5,22].AlarmTimerSP := 2, [5,22].AutoCloseTimer.ACC := 131, [5,23].Tag := 'XV024', [5,23].CloseStatus := 1, [5,23].ZSOverride := 1, [5,23].EnableCfg := 1, [5,23].StatusWord := 4, [5,23].Status := 4, [5,23].OutputAddress := 55, [5,23].AlarmTimer.PRE := 2000, [5,23].AlarmTimerSP := 2, [5,23].AutoCloseTimer.ACC := 1003, [5,24].Tag := 'XV025', [5,24].CloseStatus := 1,
        [5,24].ZSOverride := 1, [5,24].EnableCfg := 1, [5,24].StatusWord := 4, [5,24].Status := 4, [5,24].OutputAddress := 56, [5,24].AlarmTimer.PRE := 2000, [5,24].AlarmTimerSP := 2, [5,24].AutoCloseTimer.ACC := 1002, [5,25].Tag := 'XV026', [5,25].CloseStatus := 1, [5,25].ZSOverride := 1, [5,25].EnableCfg := 1, [5,25].StatusWord := 4, [5,25].Status := 4, [5,25].OutputAddress := 57, [5,25].AlarmTimer.PRE := 2000, [5,25].AlarmTimerSP := 2, [5,25].AutoCloseTimer.ACC := 1002, [5,26].Tag := 'XV028', [5,26].CloseStatus := 1, [5,26].ZSOverride := 1, [5,26].EnableCfg := 1, [5,26].StatusWord := 4, [5,26].Status := 4, [5,26].OutputAddress := 58, [5,26].AlarmTimer.PRE := 2000, [5,26].AlarmTimerSP := 2, [5,26].AutoCloseTimer.ACC := 1002, [5,27].Tag := 'XV029', [5,27].CloseStatus := 1, [5,27].ZSOverride := 1, [5,27].EnableCfg := 1, [5,27].StatusWord := 4, [5,27].Status := 4, [5,27].OutputAddress := 59, [5,27].AlarmTimer.PRE := 2000, [5,27].AlarmTimerSP := 2, [5,28].Tag := 'XV030', [5,28].CloseStatus := 1, [5,28].ZSOverride := 1, [5,28].EnableCfg := 1, [5,28].StatusWord := 4, [5,28].Status := 4, [5,28].OutputAddress := 60, [5,28].AlarmTimer.PRE := 2000, [5,28].AlarmTimerSP := 2, [5,29].Tag := 'XV031', [5,29].Control := 1, [5,29].Auto := 1, [5,29].Manual := 1, [5,29].OpenStatus := 1, [5,29].ZSOverride := 1, [5,29].FailState := 1, [5,29].EnableCfg := 1, [5,29].StatusWord := 2, [5,29].Status := 2, [5,29].OutputAddress := 61, [5,29].AlarmTimer.PRE := 2000, [5,29].AlarmTimerSP := 2, [5,29].AutoCloseTimer.ACC := 1068,
        [5,30].Tag := 'XV033', [5,30].CloseStatus := 1, [5,30].ZSOverride := 1, [5,30].EnableCfg := 1, [5,30].StatusWord := 4, [5,30].Status := 4, [5,30].OutputAddress := 62, [5,30].AlarmTimer.PRE := 2000, [5,30].AlarmTimerSP := 2, [5,30].AutoCloseTimer.ACC := 1069, [5,31].Tag := 'XV034', [5,31].CloseStatus := 1, [5,31].ZSOverride := 1, [5,31].EnableCfg := 1, [5,31].StatusWord := 4, [5,31].Status := 4, [5,31].OutputAddress := 63, [5,31].AlarmTimer.PRE := 2000, [5,31].AlarmTimerSP := 2, [5,31].AutoCloseTimer.ACC := 131, [5,32].CloseStatus := 1, [5,32].PriorityCfg := 1, [5,32].ZSOpenAddress := 32, [5,32].OutputAddress := 68, [5,32].AlarmTimer.PRE := 2000, [5,32].AlarmTimerSP := 2, [5,32].AutoCloseTimer.ACC := 1059, [5,33].OpenStatus := 1, [5,33].PriorityCfg := 1, [5,33].FailState := 1, [5,33].ZSCloseAddress := 33, [5,33].OutputAddress := 69, [5,33].AlarmTimer.PRE := 2000, [5,33].AlarmTimerSP := 2, [5,33].AutoCloseTimer.ACC := 1123, [5,34].OpenStatus := 1, [5,34].PriorityCfg := 1, [5,34].FailState := 1, [5,34].ZSCloseAddress := 34, [5,34].OutputAddress := 70, [5,34].AlarmTimer.PRE := 2000, [5,34].AlarmTimerSP := 2, [5,34].AutoCloseTimer.ACC := 1095, [5,35].OpenStatus := 1, [5,35].PriorityCfg := 1, [5,35].FailState := 1, [5,35].ZSCloseAddress := 35, [5,35].OutputAddress := 71, [5,35].AlarmTimer.PRE := 2000, [5,35].AlarmTimerSP := 2, [5,35].AutoCloseTimer.ACC := 1127, [5,36].OpenStatus := 1, [5,36].PriorityCfg := 1, [5,36].FailState := 1, [5,36].ZSCloseAddress := 36, [5,36].OutputAddress := 72, [5,36].AlarmTimer.PRE := 2000, [5,36].AlarmTimerSP := 2, [5,36].AutoCloseTimer.ACC := 1004, [5,37].CloseStatus := 1,
        [5,37].PriorityCfg := 1, [5,37].ZSOpenAddress := 37, [5,37].OutputAddress := 73, [5,37].AlarmTimer.PRE := 2000, [5,37].AlarmTimerSP := 2, [5,37].AutoCloseTimer.ACC := 1121, [5,38].CloseStatus := 1, [5,38].Priority := 1, [5,38].PriorityCfg := 1, [5,38].ZSOpenAddress := 38, [5,38].OutputAddress := 40, [5,38].AlarmTimer.PRE := 2000, [5,38].AlarmTimerSP := 2, [5,38].AutoCloseTimer.ACC := 1135, [5,39].CloseStatus := 1, [5,39].Priority := 1, [5,39].PriorityCfg := 1, [5,39].ZSOpenAddress := 39, [5,39].OutputAddress := 41, [5,39].AlarmTimer.PRE := 2000, [5,39].AlarmTimerSP := 2, [5,39].AutoCloseTimer.ACC := 1121, [5,40].CloseStatus := 1, [5,40].Priority := 1, [5,40].PriorityCfg := 1, [5,40].ZSOpenAddress := 40, [5,40].OutputAddress := 42, [5,40].AlarmTimer.PRE := 2000, [5,40].AlarmTimerSP := 2, [5,40].AutoCloseTimer.ACC := 1112, [5,41].CloseStatus := 1, [5,41].Priority := 1, [5,41].PriorityCfg := 1, [5,41].ZSOpenAddress := 41, [5,41].OutputAddress := 43, [5,41].AlarmTimer.PRE := 2000, [5,41].AlarmTimerSP := 2, [5,42].CloseStatus := 1, [5,42].Priority := 1, [5,42].PriorityCfg := 1, [5,42].ZSOpenAddress := 42, [5,42].OutputAddress := 44, [5,42].AlarmTimer.PRE := 2000, [5,42].AlarmTimerSP := 2, [5,43].CloseStatus := 1, [5,43].Priority := 1, [5,43].PriorityCfg := 1, [5,43].ZSOpenAddress := 43, [5,43].OutputAddress := 52, [5,43].AlarmTimer.PRE := 2000, [5,43].AlarmTimerSP := 2, [5,44].CloseStatus := 1, [5,44].Priority := 1, [5,44].PriorityCfg := 1, [5,44].ZSOpenAddress := 44, [5,44].OutputAddress := 53, [5,44].AlarmTimer.PRE := 2000, [5,44].AlarmTimerSP := 2, [5,45].CloseStatus := 1, [5,45].Priority := 1,
        [5,45].PriorityCfg := 1, [5,45].ZSOpenAddress := 45, [5,45].OutputAddress := 54, [5,45].AlarmTimer.PRE := 2000, [5,45].AlarmTimerSP := 2, [5,46].CloseStatus := 1, [5,46].Priority := 1, [5,46].PriorityCfg := 1, [5,46].ZSOpenAddress := 46, [5,46].OutputAddress := 55, [5,46].AlarmTimer.PRE := 2000, [5,46].AlarmTimerSP := 2, [5,47].OpenStatus := 1, [5,47].Priority := 1, [5,47].PriorityCfg := 1, [5,47].FailState := 1, [5,47].ZSCloseAddress := 47, [5,47].OutputAddress := 45, [5,47].AlarmTimer.PRE := 2000, [5,47].AlarmTimerSP := 2, [5,48].FailState := 1, [5,48].ZSCloseAddress := 48, [5,48].OutputAddress := 80, [5,49].FailState := 1, [5,49].ZSCloseAddress := 49, [5,49].OutputAddress := 81, [5,50].FailState := 1, [5,50].ZSCloseAddress := 50, [5,50].OutputAddress := 82, [5,51].OpenStatus := 1, [5,51].FailState := 1, [5,51].ZSCloseAddress := 51, [5,51].OutputAddress := 83, [5,52].OpenStatus := 1, [5,52].FailState := 1, [5,52].ZSCloseAddress := 52, [5,52].OutputAddress := 84, [5,53].CloseStatus := 1, [5,53].FailState := 1, [5,53].ZSCloseAddress := 53, [5,53].OutputAddress := 85, [5,54].CloseStatus := 1, [5,54].FailState := 1, [5,54].ZSCloseAddress := 54, [5,54].OutputAddress := 86, [5,55].CloseStatus := 1, [5,55].FailState := 1, [5,55].ZSCloseAddress := 55, [5,55].OutputAddress := 87, [5,56].CloseStatus := 1, [5,58].CloseStatus := 1, [5,59].CloseStatus := 1);
   ValveControl : ValveControl := (ValveStatus1 := 387, MaxValveNum := 32);   // Valve Control
   ValveSwInput : BOOL[64];   // Valve digital input
        [2]   // XV003 Closed Switch
        [3]   // XV004 Closed Switch
        [4]   // XV005 Closed Switch
        [5]   // XV006 Closed Switch
        [6]   // XV007 Closed Switch
   VersionLetterForDevelopment : STRING := '.c';   // Version Letter for Development
   VersionNumberForRelease : STRING := '1.01.00.01';   // Version Number for Release
   WI101 : ALIAS FOR AnalogPoint[15];
   WI101Alarm : ALIAS FOR AlarmAnalog[15];
   WI201 : ALIAS FOR AnalogPoint[1];
   WI201_SIG : ALIAS FOR DigitalPoint[96];
   WI201Alarm : ALIAS FOR AlarmAnalog[1];
   XS011 : ALIAS FOR DigitalPoint[14];
   XS012 : ALIAS FOR DigitalPoint[15];
   XV001 : ALIAS FOR Valve[0];
   XV002 : ALIAS FOR Valve[1];
   XV003 : ALIAS FOR Valve[2];
   XV004 : ALIAS FOR Valve[3];
   XV005 : ALIAS FOR Valve[4];
   XV006 : ALIAS FOR Valve[5];
   XV007 : ALIAS FOR Valve[6];
   XV101 : ALIAS FOR Valve[7];
   XV102 : ALIAS FOR Valve[8];
   XV201 : ALIAS FOR Valve[15];
   XV202 : ALIAS FOR Valve[16];
   XV401 : ALIAS FOR Valve[9];
   XV402 : ALIAS FOR Valve[10];
   XV403 : ALIAS FOR Valve[11];
   XV404 : ALIAS FOR Valve[12];
   XV405 : ALIAS FOR Valve[13];
   XV406 : ALIAS FOR Valve[14];
   XV701 : ALIAS FOR Valve[17];
   XV702 : ALIAS FOR Valve[18];
   XV703 : ALIAS FOR Valve[19];
   XV704 : ALIAS FOR Valve[20];
   Y500A : ALIAS FOR DigitalOutput[10];
   Y500B : ALIAS FOR DigitalOutput[11];
   Y501A : ALIAS FOR DigitalOutput[12];
   Y501B : ALIAS FOR DigitalOutput[13];
   YA01 : ALIAS FOR DigitalPoint[50];
   YA02 : ALIAS FOR DigitalPoint[51];
   YA03 : ALIAS FOR DigitalPoint[52];
   YA04 : ALIAS FOR DigitalPoint[53];
   YA05 : ALIAS FOR DigitalPoint[54];
   YA06 : ALIAS FOR DigitalPoint[55];
   YA07 : ALIAS FOR DigitalPoint[56];
   YA08 : ALIAS FOR DigitalPoint[57];
   YA09 : ALIAS FOR DigitalPoint[58];
   YA10 : ALIAS FOR DigitalPoint[59];
   YA11 : ALIAS FOR DigitalPoint[60];
   YA12 : ALIAS FOR DigitalPoint[61];
   YA13 : ALIAS FOR DigitalPoint[62];
   YA14 : ALIAS FOR DigitalPoint[63];
   YA15 : ALIAS FOR DigitalPoint[69];
   YA16 : ALIAS FOR DigitalPoint[70];
   YA17 : ALIAS FOR DigitalPoint[71];
   YA18 : ALIAS FOR DigitalPoint[72];
   YA41 : ALIAS FOR DigitalPoint[73];
   ZS001 : ALIAS FOR DigitalPoint[6];
   ZS002 : ALIAS FOR DigitalPoint[7];
   ZS003 : ALIAS FOR DigitalPoint[8];
   ZS004 : ALIAS FOR DigitalPoint[9];
   ZS005 : ALIAS FOR DigitalPoint[10];
   ZS008 : ALIAS FOR DigitalPoint[5];
   ZSDF : ALIAS FOR DigitalPoint[68];
END_VAR

PROGRAM CCPSystem   (* main routine MainRoutine, fault routine FaultRoutine *)
VAR
   ActionCode : DINT;   // Action Code
   ActionFlag : BOOL;   // Action Flag
   ActionProperty : DINT;   // Action Property
   ActionStructure : DINT;   // Action Data Structure
   ActionTag : DINT := 3;   // Action Tag
   ActionValue : REAL;   // Action Value
   AutoRunTimer : TIMER := (PRE := 5000);   // Auto Run Timer
   Boolean : DINT;   // Boolean Operator
        .1   // AND
        .0   // OR
   Branch : BOOL;   // Conditional Branch Flag
   BranchStep : DINT;   // Branch Step Number
   BufferStep : DINT := 3012;   // Buffer Step
   Clear : BOOL;   // Clear Operation Table Flag
   Code : DINT := 1700002;   // Global Code
   CompleteTimer : TIMER := (PRE := 10000);   // Operation Complete Timer
   Criteria1BoolValue : BOOL;   // Criteria 1 Discrete Value
   Criteria1Code : DINT := 800303;   // Criteria 1 Code
   Criteria1Met : BOOL;   // Criteria 1 Met
   Criteria1Operator : DINT := 1;   // Criteria 1 Operator
        .0   // >=
        .1   // <=
        .2   // =
   Criteria1Property : DINT := 3;   // Criteria 1 Property
   Criteria1RealValue : REAL := 2.0;   // Criteria 1 Real Value
   Criteria1Structure : DINT := 8;   // Criteria 1 Data Structure
   Criteria1Tag : DINT := 3;   // Criteria 1 Tag
   Criteria1Type : BOOL := 1;   // Criteria 1 Type 0=Real, 1=Boolean
   Criteria1Value : REAL := 1.0;   // Criteria 1 Value
   Criteria2BoolValue : BOOL := 1;   // Criteria 2 Discrete Value
   Criteria2Code : DINT;   // Criteria 2 Code
   Criteria2Met : BOOL := 1;   // Criteria 2 Met
   Criteria2Operator : DINT;   // Criteria 2 Operator
        .0   // >=
        .1   // <=
        .2   // =
   Criteria2Property : DINT := 3;   // Criteria 2 Property
   Criteria2RealValue : REAL := 17.0;   // Criteria 2 Real Value
   Criteria2Structure : DINT;   // Criteria 2 Data Structure
   Criteria2Tag : DINT;   // Criteria 2 Tag
   Criteria2Type : BOOL;   // Criteria 2 Type 0=Real, 1=Boolean
   Criteria2Value : REAL;   // Criteria 2 Value
   CriteriaMet : BOOL;   // Criteria Met
   DateTime : DINT[7] := ([0] := 2025, [1] := 10, [2] := 3, [3] := 11, [4] := 41, [5] := 40, [6] := 147549);   // Date and Time
   DownloadONS : BOOL;
   EnableStep : BOOL;   // Step Action Enabled
   ErrorCheck : BOOL;   // Error Check Flag
   ErrorCheckONS : BOOL := 1;   // Error Check One-Shot
   Index : DINT := 710;   // Index
   LastStep : DINT := 11;   // Last Step
   NextStep : DINT := 14;   // Next Step
   PendingStep : DINT := 13;   // Current Step
   Phase0StopONS : BOOL;
   PhaseClear : BOOL;   // Phase Clear
   PhaseClearNumber : DINT := 6;   // Phase Clear Number
   PhaseNumber : DINT := 6;   // Phase FOR NEXT Index
   Pointer : DINT := 249;   // Pointer
   PreRunLog : BOOL;   // Log Pre Run Set Points
   Property : DINT := 2;   // Case Property
   Run : BOOL;   // Operation Run Status
   RunONS : BOOL;   // Run Command One-Shot
   sAction : STRING10 := '800301';   // Action Code String
   sActionProperty : STRING4 := '01';   // Action Property String
   sActionStructure : STRING4 := '8';   // Action Data Structure String
   sActionTag : STRING4 := '003';   // Action Tag String
   sBufferEvents : STRING50 := '10032025,11:37:21.0,300206,1.00000000,';   // Buffer Events String
   sCode : STRING10 := '2501101';   // Global code String
   sColon : STRING4 := ':';   // Colon separator String
   sComma : STRING4 := ',';   // Comma String
   sCriteria1 : STRING10 := '800303';   // Criteria 1 Code String
   sCriteria1Property : STRING4 := '03';   // Criteria 1 Property String
   sCriteria1Structure : STRING4 := '8';   // Criteria 1 Data Structure String
   sCriteria1Tag : STRING4 := '003';   // Criteria 1 Tag String
   sCriteria2 : STRING10 := '800003';   // Criteria 2 Code String
   sCriteria2Property : STRING4 := '03';   // Criteria 2 Property String
   sCriteria2Structure : STRING4 := '8';   // Criteria 2 Data Structure String
   sCriteria2Tag : STRING4 := '000';   // Criteria 2 Tag String
   sDateTime : STRING25 := '10032025,11:41:40.1,';   // Date and Time String
   sPeriod : STRING4 := '.';   // Timer separator String
   sProperty : STRING4 := '02';   // Property String
   sStructure : STRING4 := '17';   // Structure String
   sTag : STRING4 := '000';   // Tag String
   sTemp : STRING50 := '1';   // Temp String
   Structure : DINT := 17;   // Structure code
   sZero : STRING4 := '0';   // Zero String
   Tag : DINT;   // Tag value
   TempEvents : DINT := 50;   // Temp Register
   TempSteps : DINT := 26;
   Tenths : DINT := 1;   // Thents (Date and Time management)
   ThisStep : DINT := 66;   // This Step (Error management)
   Value : REAL := 1.0;   // Temp Value
END_VAR

ROUTINE Action   (* structured text *)
// Operation Action Routine
   (* =======================================================================
   	Operation Action : Get the current action code and perform action based on information extraction
   
   	List of treatments
   		- Get current action code
   		- Extract informations based on action code
   		- Navigate through the action categories to perform action
   		- Jump to BufferSteps routine and update step numbers
   
   -----------------------------------------------------------------------------------------------------------------------------------------------------
   	History
   		2019-DEC-24 - Merck - Q. Spindler - Initial version for Candidate Release 1.00.00.00.a
   		2020-APR-14 - Merck - Q. Spindler - Modifications for Candidate Release 1.00.00.00.b
   					- Add SysControl.Zero_WI101_Cmd
   					- Add Valve.ZSOverride for valves limit switch alarms
   					- Add Gateway actions
   		2020-SEP-18 - Merck - Q. Spindler - Modifications for Candidate Release 1.00.00.00.d
   					- Add ExternalWeight and ExternalTCU actions
   		2021-NOV-23 - Merck - Q. Spindler - Modifications for Candidate Release 1.01.00.00.a
   					- Add Reset of ResponseOK, YES, and NO on prompt action
   =========================================================================*)
   
   
   (* Get current action code
   =========================================================================*)
   (*Get the pending step Action Code and Action Value from the operation array*)
   ActionCode := Operation[PhaseNumber,PendingStep].Action;
   ActionValue := Operation[PhaseNumber,PendingStep].ActionValue;
   
   (* Extract informations based on action code
   =========================================================================*)
   (*Extract the Structure, Tag and Property values from the action code. The action code is
   in the format SSTTTPP  SS is Structure Element, TTT is action TagElement i.e ControlLoop[TTT].Enable
   PP Action Property Number in secound Case below.*)
   
   IF ActionCode <> 0 THEN;
   	DTOS (ActionCode, sAction);
   	IF sAction.LEN = 7 THEN;
   		MID (sAction, 2, 1, sActionStructure);
   		MID (sAction, 3, 3, sActionTag);
   		MID (sAction, 2, 6, sActionProperty);
   	ELSIF sAction.LEN = 6 THEN;
   		MID (sAction, 1, 1, sActionStructure);
   		MID (sAction, 3, 2, sActionTag);
   		MID (sAction, 2, 5, sActionProperty);
   	ELSIF sAction.LEN = 5 THEN;
   		(* Ignore if code length is not 6 or 7 *)
   		DTOS(0,sActionStructure);
   	ELSE;
   		CCPSystem.Error := 7;
   	END_IF;
   	STOD (sActionStructure, ActionStructure);
   	STOD (sActionTag, ActionTag);
   	STOD (sActionProperty, ActionProperty);
   ELSE;
   	ActionStructure := 0;
   END_IF;
   
   (* Navigate through the action categories to perform action
   =========================================================================*)
   CASE ActionStructure OF
   	0:	; (*No Action)*)
   	1: 	CASE	ActionProperty OF (*Analog Alarms*)
   			1:	IF NOT ErrorCheck THEN; IF ActionValue = 0 THEN AlarmAnalog[ActionTag].Override := 0; ELSE AlarmAnalog[ActionTag].Override := 1; END_IF; END_IF;
   			2:	IF NOT ErrorCheck THEN; AlarmAnalog[ActionTag].LOLO := ActionValue; END_IF;
   			3:	IF NOT ErrorCheck THEN; AlarmAnalog[ActionTag].LO := ActionValue; END_IF;
   			4:	IF NOT ErrorCheck THEN; AlarmAnalog[ActionTag].HI := ActionValue; END_IF;
   			5:	IF NOT ErrorCheck THEN; AlarmAnalog[ActionTag].HIHI := ActionValue; END_IF;
   		ELSE 	CCPSystem.Error := 7;
   		END_CASE;
   	2:	CASE	ActionProperty OF (*Deviation Alarms*)
   			1:	IF NOT ErrorCheck THEN; IF ActionValue = 0 THEN AlarmDeviation[ActionTag].Override := 0; ELSE AlarmDeviation[ActionTag].Override := 1; END_IF; END_IF;
   			4:	IF NOT ErrorCheck THEN; AlarmDeviation[ActionTag].HI := ActionValue; END_IF;
   			5:	IF NOT ErrorCheck THEN; AlarmDeviation[ActionTag].HIHI := ActionValue; END_IF;
   		ELSE 	CCPSystem.Error := 7;
   		END_CASE;
   	3:	CASE	ActionProperty OF (*Digital Alarms*)
   			1:	IF NOT ErrorCheck THEN; IF ActionValue = 0 THEN DigitalPoint[ActionTag].Override := 0; ELSE DigitalPoint[ActionTag].Override := 1; END_IF; END_IF;
   		ELSE 	CCPSystem.Error := 7;
   		END_CASE;
   	5:	CASE	ActionProperty OF (*Control Loops*)
   			1:	IF NOT ErrorCheck THEN; IF ActionValue = 0 THEN ControlLoop[ActionTag].Manual := 0; ELSE ControlLoop[ActionTag].Manual := 1; END_IF; END_IF;
   			2:	IF NOT ErrorCheck THEN; IF ActionValue = 0 THEN ControlLoop[ActionTag].Auto1 := 0; ELSE ControlLoop[ActionTag].Auto1 := 1; END_IF; END_IF;
   			3:	IF NOT ErrorCheck THEN; IF ActionValue = 0 THEN ControlLoop[ActionTag].Auto2 := 0; ELSE ControlLoop[ActionTag].Auto2 := 1; END_IF; END_IF;
   			4:	IF NOT ErrorCheck THEN; IF ActionValue = 0 THEN ControlLoop[ActionTag].Auto3 := 0; ELSE ControlLoop[ActionTag].Auto3 := 1; END_IF; END_IF;
   			5:	IF NOT ErrorCheck THEN; IF ActionValue = 0 THEN ControlLoop[ActionTag].Auto4 := 0; ELSE ControlLoop[ActionTag].Auto4 := 1; END_IF; END_IF;
   			6:	IF NOT ErrorCheck THEN; ControlLoop[ActionTag].SPManual := ActionValue; END_IF;
   			7:	IF NOT ErrorCheck THEN; ControlLoop[ActionTag].SPAuto1 := ActionValue; END_IF;
   			8:	IF NOT ErrorCheck THEN; ControlLoop[ActionTag].SPAuto2 := ActionValue; END_IF;
   			9:	IF NOT ErrorCheck THEN; ControlLoop[ActionTag].SPAuto3 := ActionValue; END_IF;
   			10:	IF NOT ErrorCheck THEN; ControlLoop[ActionTag].SPAuto4 := ActionValue; END_IF;
   			11:	IF NOT ErrorCheck THEN; ControlLoop[ActionTag].RampRate := ActionValue; END_IF;
   			12:	IF NOT ErrorCheck THEN; ControlLoop[ActionTag].Deadband := ActionValue; END_IF;
   			13:	IF NOT ErrorCheck THEN; ControlLoop[ActionTag].StableTime := ActionValue; END_IF;
   			14:	IF NOT ErrorCheck THEN; ControlLoop[ActionTag].KP[0] := ActionValue; END_IF;
   			15:	IF NOT ErrorCheck THEN; ControlLoop[ActionTag].KI[0] := ActionValue; END_IF;
   			16:	IF NOT ErrorCheck THEN; ControlLoop[ActionTag].KD[0] := ActionValue; END_IF;
   			17:	IF NOT ErrorCheck THEN; ControlLoop[ActionTag].DB[0] := ActionValue; END_IF;
   			18:	IF NOT ErrorCheck THEN; ControlLoop[ActionTag].KP[1] := ActionValue; END_IF;
   			19:	IF NOT ErrorCheck THEN; ControlLoop[ActionTag].KI[1] := ActionValue; END_IF;
   			20:	IF NOT ErrorCheck THEN; ControlLoop[ActionTag].KD[1] := ActionValue; END_IF;
   			21: IF NOT ErrorCheck THEN; ControlLoop[ActionTag].DB[1] := ActionValue; END_IF;
   			22: IF NOT ErrorCheck THEN; ControlLoop[ActionTag].KP[2] := ActionValue; END_IF;
   			23:	IF NOT ErrorCheck THEN; ControlLoop[ActionTag].KI[2] := ActionValue; END_IF;
   			24:	IF NOT ErrorCheck THEN; ControlLoop[ActionTag].KD[2] := ActionValue; END_IF;
   			25:	IF NOT ErrorCheck THEN; ControlLoop[ActionTag].DB[2] := ActionValue; END_IF;
   		ELSE 	CCPSystem.Error := 7;
   		END_CASE;
   	7:	CASE	ActionProperty OF (*Phase Control*)
   			1:	IF NOT ErrorCheck THEN; IF ActionValue = 0 THEN Phase[ActionTag].Run := 0; ELSE Phase[ActionTag].Run := 1; END_IF; END_IF;
   			2:	IF NOT ErrorCheck THEN; IF ActionValue = 0 THEN Phase[ActionTag].Stop := 0; ELSE Phase[ActionTag].Stop := 1; END_IF; END_IF;
   			3:	IF NOT ErrorCheck THEN; IF ActionValue = 0 THEN Phase[ActionTag].Hold := 0; ELSE Phase[ActionTag].Hold := 1; END_IF; END_IF;
   			4:	IF NOT ErrorCheck THEN; IF ActionValue = 0 THEN Phase[ActionTag].Pause := 0; ELSE Phase[ActionTag].Pause := 1; END_IF; END_IF;
   			5:	IF NOT ErrorCheck THEN;
   				Phase[PhaseNumber].JumpPLC := 1; (*Conditional Branch*)
   				Phase[PhaseNumber].ActualStep := BranchStep;
   				END_IF;
   		ELSE 	CCPSystem.Error := 7;
   		END_CASE;
   	8:	CASE	ActionProperty OF (*Prompts*)
   			(*Prompts OK*)
   			1:	IF NOT ErrorCheck THEN;
   					(*Delay to Prompts to allow back to back*)
   					TONR(PromptTimer);
   					PromptTimer.EN := 1;
   					PromptTimer.PRE := 1000;
   					while PromptTimer.TT and Prompt[PhaseNumber].PromptOK   do;
   					end_while;
   				Prompt[PhaseNumber].PromptYesNO := 0;
   				Prompt[PhaseNumber].PromptOK := 1;
   				Prompt[PhaseNumber].ResponseOK := 0;
   				Prompt[PhaseNumber].Step := PendingStep;
   				Prompt[PhaseNumber].Flag := 1;
   				Prompt[PhaseNumber].Pending := 1;
   				Prompt[PhaseNumber].Value := ActionValue; (*PV+*)
   				END_IF;
   			(*Prompts YesNo*)
   			2:	IF NOT ErrorCheck THEN;
   					(*Delay to Prompts to allow back to back*)
   					TONR(PromptTimer);
   					PromptTimer.EN := 1;
   					PromptTimer.PRE := 1000;
   					while PromptTimer.TT and Prompt[PhaseNumber].PromptYesNO do;
   					end_while;
   				Prompt[PhaseNumber].PromptOK := 0;
   				Prompt[PhaseNumber].PromptYesNO := 1;
   				Prompt[PhaseNumber].ResponseNo := 0;
   				Prompt[PhaseNumber].ResponseYes := 0;
   				Prompt[PhaseNumber].Step := PendingStep;
   				Prompt[PhaseNumber].Flag := 1;
   				Prompt[PhaseNumber].Pending := 1;
   				END_IF;
   			3:	IF NOT ErrorCheck THEN;
   				Prompt[PhaseNumber].Flag := 1;
   				Prompt[PhaseNumber].Step := PendingStep;
   				END_IF;
   		ELSE 	CCPSystem.Error := 7;
   		END_CASE;
   	9:	CASE	ActionProperty OF (*Pumps*)
   			1:	IF NOT ErrorCheck THEN; IF ActionValue = 0 THEN Drive[ActionTag].AutoCommand := 0; ELSE Drive[ActionTag].AutoCommand := 1; END_IF; END_IF;
   			2:	IF NOT ErrorCheck THEN; IF ActionValue = 0 THEN Drive[ActionTag].Direction := 0; ELSE Drive[ActionTag].Direction := 1; END_IF; END_IF;
   		ELSE 	CCPSystem.Error := 7;
   		END_CASE;
   	10:	CASE	ActionProperty OF (*Exchange Output *)
   			1:	IF NOT ErrorCheck THEN; Exchange_OUT.AO01 := ActionValue; END_IF;
   			2:	IF NOT ErrorCheck THEN; Exchange_OUT.AO02 := ActionValue; END_IF;
   			3:	IF NOT ErrorCheck THEN; Exchange_OUT.AO03 := ActionValue; END_IF;
   			4:	IF NOT ErrorCheck THEN; Exchange_OUT.AO04 := ActionValue; END_IF;
   			5:	IF NOT ErrorCheck THEN; IF ActionValue = 0 THEN Exchange_OUT.DO01 := 0; ELSE Exchange_OUT.DO01 := 1; END_IF; END_IF;
   			6:	IF NOT ErrorCheck THEN; IF ActionValue = 0 THEN Exchange_OUT.DO02 := 0; ELSE Exchange_OUT.DO02 := 1; END_IF; END_IF;
   			7:	IF NOT ErrorCheck THEN; IF ActionValue = 0 THEN Exchange_OUT.DO03 := 0; ELSE Exchange_OUT.DO03 := 1; END_IF; END_IF;
   			8:	IF NOT ErrorCheck THEN; IF ActionValue = 0 THEN Exchange_OUT.DO04 := 0; ELSE Exchange_OUT.DO04 := 1; END_IF; END_IF;
   			9:	IF NOT ErrorCheck THEN; IF ActionValue = 0 THEN Exchange_OUT.DO05 := 0; ELSE Exchange_OUT.DO05 := 1; END_IF; END_IF;
   			10:	IF NOT ErrorCheck THEN; IF ActionValue = 0 THEN Exchange_OUT.DO06 := 0; ELSE Exchange_OUT.DO06 := 1; END_IF; END_IF;
   			11:	IF NOT ErrorCheck THEN; IF ActionValue = 0 THEN Exchange_OUT.DO07 := 0; ELSE Exchange_OUT.DO07 := 1; END_IF; END_IF;
   			12:	IF NOT ErrorCheck THEN; IF ActionValue = 0 THEN Exchange_OUT.DO08 := 0; ELSE Exchange_OUT.DO08 := 1; END_IF; END_IF;
   		ELSE 	CCPSystem.Error := 7;
   		END_CASE;
   	11:	CASE	ActionProperty OF (*Timers*)
   			3:	IF NOT ErrorCheck THEN; IF ActionValue = 0 THEN Timers[ActionTag].Enable := 0; ELSE Timers[ActionTag].Enable := 1; END_IF; END_IF;
   			4:	IF NOT ErrorCheck THEN; IF ActionValue = 0 THEN Timers[ActionTag].Reset := 0; ELSE Timers[ActionTag].Reset := 1; END_IF; END_IF;
   		ELSE 	CCPSystem.Error := 7;
   		END_CASE;
   	12:	CASE	ActionProperty OF (*Totalizers*)
   			6:	IF NOT ErrorCheck THEN; IF ActionValue = 0 THEN Totalizer[0].Enable := 0; ELSE Totalizer[0].Enable := 1; END_IF; END_IF;
   			7:	IF NOT ErrorCheck THEN; Totalizer[0].Reset := 1; END_IF;
   			8:	IF NOT ErrorCheck THEN; IF ActionValue = 0 THEN Totalizer[1].Enable := 0; ELSE Totalizer[1].Enable := 1; END_IF; END_IF;
   			9:	IF NOT ErrorCheck THEN; Totalizer[1].Reset := 1; END_IF;
   		ELSE 	CCPSystem.Error := 7;
   		END_CASE;
   	13:	CASE	ActionProperty OF (*Valves*)
   			1:	IF NOT ErrorCheck THEN; IF ActionValue = 0 THEN Valve[ActionTag].Auto := 0; ELSE Valve[ActionTag].Auto := 1; END_IF; END_IF;
   			6:	IF NOT ErrorCheck THEN; IF ActionValue = 0 THEN Valve[ActionTag].ZSOverride := 0; ELSE Valve[ActionTag].ZSOverride := 1; END_IF; END_IF;
   		ELSE 	CCPSystem.Error := 7;
   		END_CASE;
   	14:	CASE	ActionProperty OF (*Mixer*)
   			1:	IF NOT ErrorCheck THEN; IF ActionValue = 0 THEN Mixer.Mode := 0; ELSE Mixer.Mode := 1; END_IF; END_IF;
   			2:	IF NOT ErrorCheck THEN; Mixer.SPManual := ActionValue; END_IF;
   			3:	IF NOT ErrorCheck THEN; Mixer.SPAutoMin := ActionValue; END_IF;
   			4:	IF NOT ErrorCheck THEN; Mixer.SPAutoMax := ActionValue; END_IF;
   			5:	IF NOT ErrorCheck THEN; Mixer.LevelMin := ActionValue; END_IF;
   			6:	IF NOT ErrorCheck THEN; Mixer.LevelMax := ActionValue; END_IF;
   		ELSE 	CCPSystem.Error := 7;
   		END_CASE;
   	15:	CASE	ActionProperty OF (*Misc.*)
   			1:	IF NOT ErrorCheck THEN; IF ActionValue = 0 THEN MiscBOOL[ActionTag] := 0; ELSE MiscBOOL[ActionTag] := 1; END_IF; END_IF;
   			2:	IF NOT ErrorCheck THEN; MiscDINT[ActionTag] := ActionValue; END_IF;
   			3:	IF NOT ErrorCheck THEN; MiscREAL[ActionTag] := ActionValue; END_IF;
   		ELSE 	CCPSystem.Error := 7;
   		END_CASE;
   	16:	CASE	ActionProperty OF (*Alarm Control*)
   			1:	IF NOT ErrorCheck THEN; AlarmControl.EnableAllIn := 1; END_IF;
   			2:	IF NOT ErrorCheck THEN; AlarmControl.DisableAllIn := 1; END_IF;
   			6:	IF NOT ErrorCheck THEN; AlarmControl.EnableAllAnaSigIn := 1; END_IF;
   			7:	IF NOT ErrorCheck THEN; AlarmControl.DisableAllAnaSigIn := 1; END_IF;
   		ELSE 	CCPSystem.Error := 7;
   		END_CASE;
   	17:	CASE	ActionProperty OF (*Miscellaneous*)
   			1:	IF NOT ErrorCheck THEN; SysControl.DefaultIn := 1; END_IF;
   			2:	IF NOT ErrorCheck THEN; ChartMark.In := 1; END_IF;
   			3:	IF NOT ErrorCheck THEN; SysControl.AllAutoIn := 1; END_IF;
   			4:	IF NOT ErrorCheck THEN; UserTotalizerManagement.LogUserIn := 1; END_IF;
   			5:	IF NOT ErrorCheck THEN; IF ActionValue = 0 THEN UserTotalizerManagement.StartUser := 0; ELSE UserTotalizerManagement.StartUser := 1; END_IF; END_IF;
   			6:	IF NOT ErrorCheck THEN; UserTotalizerManagement.ResetUserIn:= 1; END_IF;
   			7:	IF NOT ErrorCheck THEN; SysControl.Tare_WI101_Cmd := 1; END_IF;
   			8:	IF NOT ErrorCheck THEN; SysControl.ClearTare_WI101_Cmd := 1; END_IF;
   			9:	IF NOT ErrorCheck THEN; SysControl.UV_Auto_Zero_Cmd := 1; END_IF;
   			10:	IF NOT ErrorCheck THEN; SysControl.Zero_WI101_Cmd := 1; END_IF;
   			11:	IF NOT ErrorCheck THEN; IF ActionValue = 0 THEN CCPSystem.DefaultOnComplete := 0; ELSE CCPSystem.DefaultOnComplete := 1; END_IF; END_IF;
   			12:	IF NOT ErrorCheck THEN; UserAlarm.NonCritical1 := 1; END_IF;
   			13:	IF NOT ErrorCheck THEN; UserAlarm.Critical1 := 1; END_IF;
   			14:	IF NOT ErrorCheck THEN; UserAlarm.NonCritical2 := 1; END_IF;
   			15:	IF NOT ErrorCheck THEN; UserAlarm.Critical2 := 1; END_IF;
   			16:	IF NOT ErrorCheck THEN; SysControl.Tare_PI001_Cmd := 1; END_IF;
   			17:	IF NOT ErrorCheck THEN; SysControl.Tare_PI101_Cmd := 1; END_IF;
   			18:	IF NOT ErrorCheck THEN; SysControl.Tare_PI201_Cmd := 1; END_IF;
   			19:	IF NOT ErrorCheck THEN; SysControl.Tare_PI401_Cmd := 1; END_IF;
   			20:	IF NOT ErrorCheck THEN; SysControl.Tare_PI601_Cmd := 1; END_IF;
   			21:	IF NOT ErrorCheck THEN; IF ActionValue = 0 THEN BagInflate.cmd := 0; ELSE BagInflate.cmd := 1; END_IF; END_IF;
   			22:	IF NOT ErrorCheck THEN; IF ActionValue = 0 THEN ExternalTCU := 0; ELSE ExternalTCU := 1; END_IF; END_IF;
   			23:	IF NOT ErrorCheck THEN; IF ActionValue = 0 THEN ExternalWeight := 0; ELSE ExternalWeight := 1; END_IF; END_IF;
   		ELSE 	CCPSystem.Error := 7;
   		END_CASE;
   	18:	CASE	ActionProperty OF (*Criteria Flag*)
   			1:	IF NOT ErrorCheck THEN; IF ActionValue = 0 THEN CriteriaFlag.Flag1 := 0; ELSE CriteriaFlag.Flag1 := 1; END_IF; END_IF;
   			2:	IF NOT ErrorCheck THEN; IF ActionValue = 0 THEN CriteriaFlag.Flag2 := 0; ELSE CriteriaFlag.Flag2 := 1; END_IF; END_IF;
   			3:	IF NOT ErrorCheck THEN; IF ActionValue = 0 THEN CriteriaFlag.Flag3 := 0; ELSE CriteriaFlag.Flag3 := 1; END_IF; END_IF;
   			4:	IF NOT ErrorCheck THEN; IF ActionValue = 0 THEN CriteriaFlag.Flag4 := 0; ELSE CriteriaFlag.Flag4 := 1; END_IF; END_IF;
   			5:	IF NOT ErrorCheck THEN; IF ActionValue = 0 THEN CriteriaFlag.Flag5 := 0; ELSE CriteriaFlag.Flag5 := 1; END_IF; END_IF;
   		ELSE 	CCPSystem.Error := 7;
   		END_CASE;
   	19:	CASE	ActionProperty OF (*Concentration*)
   			1:	IF NOT ErrorCheck THEN; IF ActionValue = 0 THEN FQ_Conc.Enable := 0; ELSE FQ_Conc.Enable := 1; END_IF; END_IF;
   			2:	IF NOT ErrorCheck THEN; FQ_Conc.Reset:= 1; END_IF;
   			3:	IF NOT ErrorCheck THEN; Concentration.LogConcIn := 1; END_IF;
   			4:	IF NOT ErrorCheck THEN; Concentration.Conc_Init := ActionValue; END_IF;
   			5:	IF NOT ErrorCheck THEN; Concentration.Conc_Final := ActionValue; END_IF;
   			6:	IF NOT ErrorCheck THEN; Concentration.Conc_Final_Volume := ActionValue; END_IF;
   			7:	IF NOT ErrorCheck THEN; DerivedData.HOLDUP := ActionValue; END_IF;
   		ELSE 	CCPSystem.Error := 7;
   		END_CASE;
   	20:	CASE	ActionProperty OF (*Diafiltration*)
   			1:	IF NOT ErrorCheck THEN; IF ActionValue = 0 THEN FQ_Diaf.Enable := 0; ELSE FQ_Diaf.Enable := 1; END_IF; END_IF;
   			2:	IF NOT ErrorCheck THEN; FQ_Diaf.Reset:= 1; END_IF;
   			3:	IF NOT ErrorCheck THEN; Diafiltration.LogDiafIn := 1; END_IF;
   			4:	IF NOT ErrorCheck THEN; Diafiltration.Snap := 1; END_IF;
   			5:	IF NOT ErrorCheck THEN; Diafiltration.Diaf_Init := ActionValue; END_IF;
   			6:	IF NOT ErrorCheck THEN; Diafiltration.Diaf_Final_Volume := ActionValue; END_IF;
   		ELSE 	CCPSystem.Error := 7;
   		END_CASE;
   	21:	CASE	ActionProperty OF (*Membrane Data*)
   			1:	IF NOT ErrorCheck THEN; Membrane_Data.Area := ActionValue; END_IF;
   			2:	IF NOT ErrorCheck THEN; Membrane_Data.Density := ActionValue; END_IF;
   		ELSE 	CCPSystem.Error := 7;
   		END_CASE;
   	22:	CASE	ActionProperty OF (*Gateway*)
   			(*Digital Actions*)
   			1:	IF ActionTag <=31 THEN;
   					IF NOT ErrorCheck THEN; IF ActionValue = 0 THEN Gateway.RecipeAction_Digital[0].[ActionTag]:= 0; ELSE Gateway.RecipeAction_Digital[0].[ActionTag]:= 1; END_IF; END_IF;
   				ELSIF ActionTag <=63 THEN;
   					IF NOT ErrorCheck THEN; IF ActionValue = 0 THEN Gateway.RecipeAction_Digital[1].[ActionTag-32]:= 0; ELSE Gateway.RecipeAction_Digital[1].[ActionTag-32]:= 1; END_IF; END_IF;
   				END_IF;
   			(*Analog Actions*)
   			2:	IF ActionTag <=19 THEN;
   					IF NOT ErrorCheck THEN;  Gateway.RecipeAction_Analog[ActionTag] := ActionValue; END_IF;
   				END_IF;
   		ELSE 	CCPSystem.Error := 7;
   		END_CASE;
   	23:	CASE	ActionProperty OF (*PCV Control*)
   			1:	IF NOT ErrorCheck THEN; PCV101_Control.FullOpen := 1; END_IF;
   			2:	IF NOT ErrorCheck THEN; PCV101_Control.FullClose := 1; END_IF;
   			3:	IF NOT ErrorCheck THEN; PCV201_Control.FullOpen := 1; END_IF;
   			4:	IF NOT ErrorCheck THEN; PCV201_Control.FullClose := 1; END_IF;
   		ELSE 	CCPSystem.Error := 7;
   		END_CASE;
   	24:	CASE	Property OF (*Event value.*)
   			1:	IF NOT ErrorCheck THEN; LogVal.Value[Tag] := ActionValue; END_IF;
   		ELSE 	CCPSystem.Error := 7;
   		END_CASE;
   	25:	CASE	ActionProperty OF (*Flow Paths*)
   			1:	IF NOT ErrorCheck THEN; IF ActionValue = 0 THEN FlowPath[ActionTag].Command := 0; ELSE FlowPath[ActionTag].Command := 1; END_IF; END_IF;
   		ELSE 	CCPSystem.Error := 7;
   		END_CASE;
   	26:	CASE	ActionProperty OF (*Clamshell*)
   			1:	IF NOT ErrorCheck THEN; IF ActionValue = 0 THEN Y500A := 0; ELSE Y500A := 1; END_IF; END_IF;
   			2:	IF NOT ErrorCheck THEN; IF ActionValue = 0 THEN Y500B := 0; ELSE Y500B := 1; END_IF; END_IF;
   			3:	IF NOT ErrorCheck THEN; IF ActionValue = 0 THEN Y501A := 0; ELSE Y501A := 1; END_IF; END_IF;
   			4:	IF NOT ErrorCheck THEN; IF ActionValue = 0 THEN Y501B := 0; ELSE Y501B := 1; END_IF; END_IF;
   		ELSE 	CCPSystem.Error := 7;
   		END_CASE;
   	27:	CASE	ActionProperty OF (*TIC*)
   			1:	IF NOT ErrorCheck THEN; IF ActionValue = 0 THEN TIC101Control.AutoCommand := 0; ELSE TIC101Control.AutoCommand := 1; END_IF; END_IF;
   			3:	IF NOT ErrorCheck THEN; TIC101Control.Offset := ActionValue; END_IF;
   			4:	IF NOT ErrorCheck THEN; TIC101Control.OffsetTime := ActionValue; END_IF;
   			5:	IF NOT ErrorCheck THEN; TIC101Control.LevelMin := ActionValue; END_IF;
   		ELSE 	CCPSystem.Error := 7;
   		END_CASE;
   ELSE 	CCPSystem.Error := 7;
   END_CASE;
   
   
   (* Jump to BufferSteps routine and update step numbers
   =========================================================================*)
   IF NOT ErrorCheck THEN;
   	JSR (BufferSteps);
   	IF NOT Phase[PhaseNumber].JumpPLC THEN;
   		(*Update Actual step, pending step and jump step number*)
   		Phase[PhaseNumber].ActualStep := PendingStep + 1;
   		PendingStep := PendingStep + 1;
   		Phase[PhaseNumber].JumpStep := PendingStep + 1;
   	END_IF;
   END_IF;
END_ROUTINE
